// TIA Portal V20 export
Screen "SafetyZone06Overview"  1276x673
  ScreenItem "Button_Overview_LegendᆉY2" at 1185,2 size 90x60  Type=HmiButton
  ScreenItem "Button_Back" at 2,4 size 90x60  Type=HmiButton
  ScreenItem "Rectangle_12" at 202,545 size 726x8  Type=HmiRectangle
  ScreenItem "Line_Header_X0_Y64" at -11,64 size 1280x0  Type=HmiLine
  ScreenItem "Emerg_2" at 264,552 size 52x56  Type=HmiSymbolicIOField
  ScreenItem "Graphic view_19" at 833,324 size 46x35  Type=HmiGraphicView
  ScreenItem "Faceplate container_2" at 347,404 size 104x136  Type=HmiFaceplateContainer
  ScreenItem "Faceplate container_11" at 469,274 size 362x136  Type=HmiFaceplateContainer
  ScreenItem "Faceplate container_16" at 873,298 size 152x87  Type=HmiFaceplateContainer
  ScreenItem "Faceplate container_17" at 689,556 size 152x87  Type=HmiFaceplateContainer
  ScreenItem "Faceplate container_18" at 496,556 size 152x87  Type=HmiFaceplateContainer
  ScreenItem "Faceplate container_6" at 467,405 size 110x138  Type=HmiFaceplateContainer
  ScreenItem "Faceplate container_1" at 815,405 size 110x140  Type=HmiFaceplateContainer
  ScreenItem "Rectangle_6" at 202,125 size 724x8  Type=HmiRectangle
  ScreenItem "Rectangle_7" at 954,202 size 160x8  Type=HmiRectangle
  ScreenItem "Rectangle_11" at 954,462 size 160x8  Type=HmiRectangle
  ScreenItem "Rectangle_14" at 127,202 size 160x8  Type=HmiRectangle
  ScreenItem "Rectangle_15" at 127,462 size 160x8  Type=HmiRectangle
  ScreenItem "Rectangle_16" at 272,595 size 88x8  Type=HmiRectangle
  ScreenItem "Rectangle_17" at 434,594 size 88x8  Type=HmiRectangle
  ScreenItem "Faceplate container_22" at 636,131 size 110x145  Type=HmiFaceplateContainer
  ScreenItem "Graphic view_2" at 248,591 size 77x60  Type=HmiGraphicView
  ScreenItem "Faceplate container_8" at 699,405 size 110x147  Type=HmiFaceplateContainer
  ScreenItem "Graphic view_4" at 312,324 size 46x35  Type=HmiGraphicView
  ScreenItem "Faceplate container_23" at 809,134 size 110x140  Type=HmiFaceplateContainer
  ScreenItem "图形 IO 域_26" at 202,271 size 15x122  Type=HmiSymbolicIOField
  ScreenItem "图形 IO 域_15" at 1027,271 size 15x122  Type=HmiSymbolicIOField
  ScreenItem "图形 IO 域_16" at 391,578 size 15x119  Type=HmiSymbolicIOField
  ScreenItem "图形 IO 域_17" at 456,554 size 15x90  Type=HmiSymbolicIOField
  ScreenItem "图形 IO 域_18" at 325,553 size 15x90  Type=HmiSymbolicIOField
  ScreenItem "Button_Overview_LegendᆉY2_1" at 1092,2 size 90x60  Type=HmiButton
  ScreenItem "文本域_2" at 981,601 size 58x19  Type=HmiTextBox
  ScreenItem "矩形_1" at 928,543 size 14x11  Type=HmiRectangle
  ScreenItem "线_1" at 941,558 size 47x13  Type=HmiLine
  ScreenItem "矩形_2" at 941,543 size 48x11  Type=HmiRectangle
  ScreenItem "矩形_3" at 988,543 size 14x11  Type=HmiRectangle
  ScreenItem "Button_Overview_LegendᆉY2_2" at 986,2 size 103x60  Type=HmiButton
  ScreenItem "Rectangle_30" at 1002,545 size 36x8  Type=HmiRectangle
  ScreenItem "Title_ScreenOverview_X390_Y2_1" at 384,4 size 510x57  Type=HmiTextBox
  ScreenItem "Button_Overview_LegendᆉY2_3" at 106,2 size 103x60  Type=HmiButton
  ScreenItem "Faceplate container_3" at 581,405 size 110x147  Type=HmiFaceplateContainer
  ScreenItem "文本域_3" at 844,560 size 50x20  Type=HmiTextBox
  ScreenItem "Emerg_6" at 841,573 size 52x56  Type=HmiSymbolicIOField
  ScreenItem "Fusszeile_Button_ManualOPMode1_4" at 246,404 size 90x60  Type=HmiButton
  ScreenItem "Fusszeile_Button_ManualOPMode1_3" at 246,476 size 90x60  Type=HmiButton
  ScreenItem "Faceplate container_4" at 471,135 size 110x140  Type=HmiFaceplateContainer
  ScreenItem "Emerg_1" at 975,555 size 52x56  Type=HmiSymbolicIOField
  ScreenItem "文本域_1" at 980,181 size 58x19  Type=HmiTextBox
  ScreenItem "矩形_4" at 928,123 size 14x11  Type=HmiRectangle
  ScreenItem "线_2" at 941,138 size 47x13  Type=HmiLine
  ScreenItem "矩形_5" at 941,123 size 48x11  Type=HmiRectangle
  ScreenItem "矩形_6" at 988,123 size 14x11  Type=HmiRectangle
  ScreenItem "Rectangle_1" at 1002,125 size 36x8  Type=HmiRectangle
  ScreenItem "Emerg_3" at 975,135 size 52x56  Type=HmiSymbolicIOField
